Fanuc KAREL source: kc00038.KL

-- PROVISIONAL review KL for V770-1; original PC SHA256 1fdace6419e3186fd1629f7f0ae7f6de06d9ea8ce453b07e6488c1f99575c794
-- Incomplete behavior may be omitted. Consult companion uncertainty JSON. Do not deploy.
PROGRAM KC00038
%NOLOCKGROUP
BEGIN
  -- UNRESOLVED_PC offsets 5-32; opcodes 27,22,1C,22,22,76
  -- UNRESOLVED_PC offsets 37-41; opcodes 7F
END KC00038
